FUNCTION_BLOCK SKILL_NoEquipment (* Stands in for the equipment of a primitive that has none (one that only waits): plays every command at once. Technical: Stands in for the equipment of a primitive that has none: answers every SEND with PLAYED at once *)
  (* Standard: 61499-2 *)
  (* Version 0.1, 2026-09-28, Project contributors, AAU Smart Production Lab *)
  PACKAGE modlib;
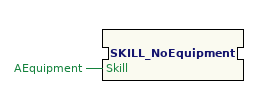
  SOCKETS
    Skill : modlib::AEquipment; (* The run's commands (AEquipment): each is played at once *)
  END_SOCKETS
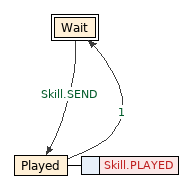
  EC_STATES
    Wait;
    Played : -> Skill.PLAYED;
  END_STATES
  EC_TRANSITIONS
    Wait TO Played := Skill.SEND;
    Played TO Wait := 1;
  END_TRANSITIONS
END_FUNCTION_BLOCK
